// TIA Portal V19 program export: 1 tag tables, 1 data types, 1 data blocks, 3 code blocks (in call order from the OBs), 0 instance data blocks

VAR_GLOBAL   // PLC tag table "Example_Tags"
   Example_Run AT %I0.0 : Bool;   // Run request
   Example_MotorOn AT %Q0.0 : Bool;
   Example_Speed AT %IW64 : Int;
END_VAR
VAR_GLOBAL CONSTANT   // user constants
   Example_MaxSpeed : Int := 1500;
END_VAR

TYPE "UDT_ExampleCfg"
   STRUCT
      Enable : Bool;
      Delay : Time := T#5S;
   END_STRUCT;
END_TYPE

DATA_BLOCK "DB_ExampleData"   // DB1
{ S7_Optimized_Access := 'TRUE' }
// stored: IsOnlyStoredInLoadMemory false, IsWriteProtectedInAS false
   VAR
      Speed : Real := 0.0;
      Scaled : Int;
   END_VAR
   VAR RETAIN
      Limit { S7_SetPoint := 'True'} : Real := 90.0;   // High speed limit
   END_VAR
   VAR
      Cfg : Struct
         Enable : Bool := true;
         Delay : Time := T#5S;
      END_STRUCT;
      Steps : Array[0..1] of Int;
   END_VAR
BEGIN
   Steps[0] := 10;
   Steps[1] := 20;
END_DATA_BLOCK

ORGANIZATION_BLOCK "Main"   // OB1, LAD, Example_ProgramCycle
// stored: AutoNumber false, IsKnowHowProtected false, ModifiedDate 2026-01-10T09:00:00.0000000Z, PriorityNumber 1
   VAR_INPUT
      Initial_Call : Bool;
   END_VAR
BEGIN

REGION Network 1: Run permissive
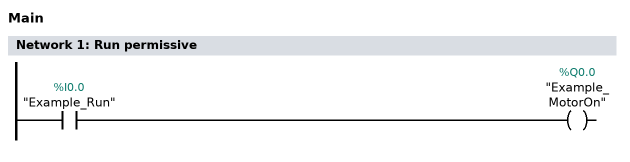
   RUNG wire#powerrail
      Contact( "Example_Run" )
      Coil( "Example_MotorOn" )
   END_RUNG
   // the same network as SCL:
   "Example_MotorOn" := "Example_Run";
END_REGION

REGION Network 2 (SCL): Speed handling
   "DB_ExampleData".Speed := "Example_Speed";
   "FC_ExampleScale"(In := "Example_Speed", Out => "DB_ExampleData".Scaled);
END_REGION
END_ORGANIZATION_BLOCK

FUNCTION "FC_ExampleScale" : Void   // FC20, STL
// stored: IsKnowHowProtected false
   VAR_INPUT
      In : Int;
   END_VAR
   VAR_OUTPUT
      Out : Int;
   END_VAR
BEGIN

NETWORK
TITLE = 
      L     #In;
      L     10;
      *I;
      T     #Out;

//scaled by ten
END_FUNCTION

FUNCTION_BLOCK "FB_ExampleValve"   // FB10, SCL
{ S7_Optimized_Access := 'TRUE' }
VERSION : 0.1
// Example valve block (synthetic)
// stored: AutoNumber true, CodeModifiedDate 2026-01-10T09:00:00.0000000Z, CompileDate 2026-01-10T09:05:00.0000000Z, IsConsistent true, IsIECCheckEnabled false, IsKnowHowProtected false, ModifiedDate 2026-01-10T09:00:00.0000000Z, SetENOAutomatically false
   VAR_INPUT
      Open : Bool;   // Open command
      Interlock : Bool;
   END_VAR
   VAR_OUTPUT
      Output : Bool;
   END_VAR
   VAR RETAIN
      OpenCount : DInt := 0;
   END_VAR
   VAR
      Limit : Real := 90.0;
   END_VAR
   VAR CONSTANT
      MaxCount : DInt := 1000;
   END_VAR
BEGIN
// Valve logic
   // Example valve permissive
   IF #Open AND NOT #Interlock THEN
       #Output := TRUE;
       #OpenCount := #OpenCount + 1; (*count openings*)
   ELSE
       #Output := FALSE;
   END_IF;
END_FUNCTION_BLOCK
